FUNCTION_BLOCK PUMP_ROTATION (* Migrated from IEC 61131-3 ST *)
  (* Standard: 61499-2 *)
  (* Version 1.0, 2026-11-06, st2fb *)
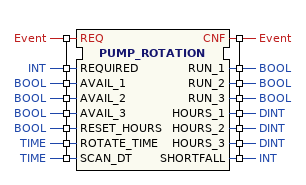
  EVENT_INPUT
    REQ WITH REQUIRED, AVAIL_1, AVAIL_2, AVAIL_3, RESET_HOURS, ROTATE_TIME, SCAN_DT;
  END_EVENT
  EVENT_OUTPUT
    CNF WITH RUN_1, RUN_2, RUN_3, HOURS_1, HOURS_2, HOURS_3, SHORTFALL;
  END_EVENT
  VAR_INPUT
    REQUIRED : INT;
    AVAIL_1 : BOOL;
    AVAIL_2 : BOOL;
    AVAIL_3 : BOOL;
    RESET_HOURS : BOOL;
    ROTATE_TIME : TIME;
    SCAN_DT : TIME;
  END_VAR
  VAR_OUTPUT
    RUN_1 : BOOL;
    RUN_2 : BOOL;
    RUN_3 : BOOL;
    HOURS_1 : DINT;
    HOURS_2 : DINT;
    HOURS_3 : DINT;
    SHORTFALL : INT;
  END_VAR
  VAR
    ST2FB_NOW : TIME := T#0s;
    ROTATE_TIMER_IN : BOOL;
    ROTATE_TIMER_PT : TIME;
    ROTATE_TIMER_Q : BOOL;
    ROTATE_TIMER_ET : TIME;
    ROTATE_TIMER_STATE : INT;
    ROTATE_TIMER_PREV_IN : BOOL;
    ROTATE_TIMER_START_TIME : TIME;
    PREV_REQUIRED : INT;
    PREV_AVAIL_1 : BOOL;
    PREV_AVAIL_2 : BOOL;
    PREV_AVAIL_3 : BOOL;
    N : INT;
    P : INT;
    BEST : INT;
    BEST_HOURS : DINT;
    CANDIDATE : BOOL;
    CANDIDATE_HOURS : DINT;
  END_VAR
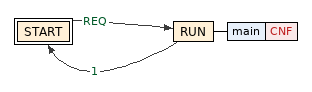
  EC_STATES
    START;
    RUN : main -> CNF;
  END_STATES
  EC_TRANSITIONS
    START TO RUN := REQ;
    RUN TO START := 1;
  END_TRANSITIONS
  ALGORITHM main IN ST:
ST2FB_NOW := ST2FB_NOW + SCAN_DT;
ROTATE_TIMER_IN := NOT ROTATE_TIMER_Q;
ROTATE_TIMER_PT := ROTATE_TIME;
IF (ROTATE_TIMER_STATE = 0) AND NOT ROTATE_TIMER_PREV_IN AND ROTATE_TIMER_IN THEN
  ROTATE_TIMER_STATE := 1;
  ROTATE_TIMER_Q := FALSE;
  ROTATE_TIMER_START_TIME := ST2FB_NOW;
ELSE
  IF NOT ROTATE_TIMER_IN THEN
    ROTATE_TIMER_ET := T#0s;
    ROTATE_TIMER_Q := FALSE;
    ROTATE_TIMER_STATE := 0;
  ELSIF ROTATE_TIMER_STATE = 1 THEN
    IF ROTATE_TIMER_START_TIME + ROTATE_TIMER_PT <= ST2FB_NOW THEN
      ROTATE_TIMER_STATE := 2;
      ROTATE_TIMER_Q := TRUE;
      ROTATE_TIMER_ET := ROTATE_TIMER_PT;
    ELSE
      ROTATE_TIMER_ET := ST2FB_NOW - ROTATE_TIMER_START_TIME;
    END_IF;
  END_IF;
END_IF;
ROTATE_TIMER_PREV_IN := ROTATE_TIMER_IN;
IF ROTATE_TIMER_Q OR (REQUIRED <> PREV_REQUIRED)
   OR (AVAIL_1 XOR PREV_AVAIL_1) OR (AVAIL_2 XOR PREV_AVAIL_2) OR (AVAIL_3 XOR PREV_AVAIL_3) THEN
  RUN_1 := FALSE;
  RUN_2 := FALSE;
  RUN_3 := FALSE;
  SHORTFALL := 0;
  FOR N := 1 TO REQUIRED DO
    BEST := 0;
    BEST_HOURS := 2147483647;
    FOR P := 1 TO 3 DO
      CASE P OF
        1:
          CANDIDATE := AVAIL_1 AND NOT RUN_1;
          CANDIDATE_HOURS := HOURS_1;
        2:
          CANDIDATE := AVAIL_2 AND NOT RUN_2;
          CANDIDATE_HOURS := HOURS_2;
        3:
          CANDIDATE := AVAIL_3 AND NOT RUN_3;
          CANDIDATE_HOURS := HOURS_3;
      END_CASE;
      IF CANDIDATE AND CANDIDATE_HOURS < BEST_HOURS THEN
        BEST := P;
        BEST_HOURS := CANDIDATE_HOURS;
      END_IF;
    END_FOR;
    CASE BEST OF
      0:
        SHORTFALL := SHORTFALL + 1;
      1:
        RUN_1 := TRUE;
      2:
        RUN_2 := TRUE;
      3:
        RUN_3 := TRUE;
    END_CASE;
  END_FOR;
END_IF;
PREV_REQUIRED := REQUIRED;
PREV_AVAIL_1 := AVAIL_1;
PREV_AVAIL_2 := AVAIL_2;
PREV_AVAIL_3 := AVAIL_3;
IF RESET_HOURS THEN
  HOURS_1 := 0;
  HOURS_2 := 0;
  HOURS_3 := 0;
ELSE
  IF RUN_1 THEN
    HOURS_1 := HOURS_1 + 1;
  END_IF;
  IF RUN_2 THEN
    HOURS_2 := HOURS_2 + 1;
  END_IF;
  IF RUN_3 THEN
    HOURS_3 := HOURS_3 + 1;
  END_IF;
END_IF;
  END_ALGORITHM
END_FUNCTION_BLOCK
(* other elements stored in the file *)
(* VarDeclaration Name=ST2FB_NOW Type=TIME InitialValue=T#0s *)
(* VarDeclaration Name=ROTATE_TIMER_IN Type=BOOL *)
(* VarDeclaration Name=ROTATE_TIMER_PT Type=TIME *)
(* VarDeclaration Name=ROTATE_TIMER_Q Type=BOOL *)
(* VarDeclaration Name=ROTATE_TIMER_ET Type=TIME *)
(* VarDeclaration Name=ROTATE_TIMER_STATE Type=INT *)
(* VarDeclaration Name=ROTATE_TIMER_PREV_IN Type=BOOL *)
(* VarDeclaration Name=ROTATE_TIMER_START_TIME Type=TIME *)
(* VarDeclaration Name=PREV_REQUIRED Type=INT *)
(* VarDeclaration Name=PREV_AVAIL_1 Type=BOOL *)
(* VarDeclaration Name=PREV_AVAIL_2 Type=BOOL *)
(* VarDeclaration Name=PREV_AVAIL_3 Type=BOOL *)
(* VarDeclaration Name=N Type=INT *)
(* VarDeclaration Name=P Type=INT *)
(* VarDeclaration Name=BEST Type=INT *)
(* VarDeclaration Name=BEST_HOURS Type=DINT *)
(* VarDeclaration Name=CANDIDATE Type=BOOL *)
(* VarDeclaration Name=CANDIDATE_HOURS Type=DINT *)
